FUNCTION_BLOCK FB_PendantState IMPLEMENTS I_PendantState
VAR
	TxBuffer	: ComBuffer;
	RxBuffer	: ComBuffer;
	pPendant : POINTER TO FB_PendantControl;
END_VAR

{warning 'add method implementation '}
METHOD DecCommand : BOOL
END_METHOD

METHOD FB_init : BOOL
VAR_INPUT
	bInitRetains : BOOL; // if TRUE, the retain variables are initialized (warm start / cold start)
	bInCopyCode : BOOL;  // if TRUE, the instance afterwards gets moved into the copy code (online change)
	pPendant : POINTER TO FB_PendantControl;

END_VAR
THIS^.pPendant := pPendant;
END_METHOD

{warning 'add method implementation '}
METHOD FocusCommand : BOOL
END_METHOD

{warning 'add method implementation '}
METHOD FoundError : BOOL
END_METHOD

{warning 'add method implementation '}
METHOD HaCommand : BOOL
END_METHOD

{warning 'add method implementation '}
METHOD InitCommand : BOOL
END_METHOD

{warning 'add method implementation '}
METHOD ResetCommand : BOOL
END_METHOD

{warning 'add method implementation '}
METHOD RunState : BOOL
END_METHOD

{warning 'add property implementation'}
PROPERTY StateID : STRING
GET
END_GET
END_PROPERTY

{warning 'add method implementation '}
METHOD Timeout : BOOL
END_METHOD

{warning 'add method implementation '}
METHOD ToIdle : BOOL
END_METHOD

END_FUNCTION_BLOCK

(* stored: Version 1.1.0.1, ProductVersion 3.1.4024.15
   POU FB_PendantState: Id {4ca28e58-094a-444e-8b9c-2a876dbabf16}, SpecialFunc None
   Method DecCommand: Id {5b2faf71-9741-463b-83a8-3063229cc9ff}
   Method FB_init: Id {fbf1ccc4-aa4d-4835-962d-1069f0a71de5}
   Method FocusCommand: Id {81666930-4619-4197-a86b-ac77eb31ce1e}
   Method FoundError: Id {35b9bb04-fbd7-46bb-ac85-34445fbee5e1}
   Method HaCommand: Id {9a83f246-765c-4cbd-9f40-7b8d8c39291a}
   Method InitCommand: Id {978c8311-d3eb-4e7f-ac97-a2d3aeaf08e4}
   Method ResetCommand: Id {9ad5f9a4-aa1c-4b5c-a9c0-c33b96b650cb}
   Method RunState: Id {f0180414-0077-4cfb-b665-58b806ee4a9b}
   Property StateID: Id {d361953c-6f62-4e53-98ce-e0644fb0ff64}
   Get Get: Id {2c15184f-f972-4d7c-a748-8085ac44079d}
   Method Timeout: Id {537e26eb-05b6-4336-83f1-89c2b678563c}
   Method ToIdle: Id {9100f539-d4ca-4611-8ce4-9948515f758a} *)
